(* IEC 61131-3 sources: model-first-plc-agent-ai/results/T3-W-09, 2 files *)

(* ---- a1_code.st ---- *)
FUNCTION_BLOCK TankSequence
VAR_INPUT
    start : BOOL;
    stop : BOOL;
    LSH : BOOL;
    LSHH : BOOL;
    TON_Duration : TIME;
    TOF_Duration : TIME;
END_VAR
VAR_OUTPUT
    fill_valve : BOOL;
    discharge_valve : BOOL;
END_VAR
VAR
    active_state : INT := 0;
    filling_active : BOOL;
    ton_q : BOOL;
    tof_q : BOOL;
    fill_timer : TON;
    pause_timer : TOF;
END_VAR

(* Evaluate both timers every scan using the current filling-step activity. *)
filling_active := (active_state = 1);

fill_timer(IN := filling_active, PT := TON_Duration);
pause_timer(IN := filling_active, PT := TOF_Duration);

ton_q := fill_timer.Q;
tof_q := pause_timer.Q;

(* Evaluate transitions from the current situation only. *)
CASE active_state OF
    0:
        IF start AND NOT stop AND NOT LSH AND NOT LSHH THEN
            active_state := 1;
        END_IF;

    1:
        IF stop OR LSH OR LSHH THEN
            active_state := 0;
        ELSIF ton_q AND NOT stop AND NOT LSH AND NOT LSHH THEN
            active_state := 2;
        END_IF;

    2:
        IF stop OR LSH OR LSHH THEN
            active_state := 0;
        ELSIF NOT tof_q AND NOT stop AND NOT LSH AND NOT LSHH THEN
            active_state := 1;
        END_IF;

ELSE
    active_state := 0;
END_CASE;

(* Continuous actions of the resulting situation. *)
fill_valve := (active_state = 1);
discharge_valve := FALSE;

END_FUNCTION_BLOCK

PROGRAM Main
VAR
    StartCommand AT %IX100.0 : BOOL;
    StopCommand AT %IX100.1 : BOOL;
    LSH AT %IX100.2 : BOOL;
    LSHH AT %IX100.3 : BOOL;
    FillValve AT %QX100.0 : BOOL;
    DischargeValve AT %QX100.1 : BOOL;
END_VAR
VAR
    (* Configurable example presets. *)
    TON_Duration : TIME := T#5s;
    TOF_Duration : TIME := T#5s;
    initialized : BOOL := FALSE;
    start : BOOL := FALSE;
    start_edge : R_TRIG;
    sequence_runtime : TankSequence;
END_VAR

IF NOT initialized THEN
    FillValve := FALSE;
    DischargeValve := FALSE;
    initialized := TRUE;
END_IF;

start_edge(CLK := StartCommand);
start := start_edge.Q;

sequence_runtime(
    start := start,
    stop := StopCommand,
    LSH := LSH,
    LSHH := LSHH,
    TON_Duration := TON_Duration,
    TOF_Duration := TOF_Duration
);

FillValve := sequence_runtime.fill_valve;
DischargeValve := sequence_runtime.discharge_valve;

END_PROGRAM

(* ---- a2_code.st ---- *)
FUNCTION_BLOCK TankFillingControl
VAR_INPUT
    StartCommand : BOOL;
    StopCommand : BOOL;
    LSH : BOOL;
    LSHH : BOOL;
    TON_Duration : TIME;
    TOF_Duration : TIME;
END_VAR
VAR_OUTPUT
    fill_valve : BOOL;
    discharge_valve : BOOL;
END_VAR
VAR
    ActiveState : INT := 0;
    StartEdge : R_TRIG;
    FillingTimer : TON;
    PauseTimer : TOF;
    start : BOOL;
    stop : BOOL;
    ton_q : BOOL;
    tof_q : BOOL;
    FillingActive : BOOL;
END_VAR

StartEdge(CLK := StartCommand);
start := StartEdge.Q;
stop := StopCommand;

FillingActive := (ActiveState = 1);

FillingTimer(
    IN := FillingActive,
    PT := TON_Duration
);

PauseTimer(
    IN := FillingActive,
    PT := TOF_Duration
);

ton_q := FillingTimer.Q;
tof_q := PauseTimer.Q;

IF stop THEN
    ActiveState := 0;
ELSE
    CASE ActiveState OF
        0:
            IF start AND NOT LSH THEN
                ActiveState := 1;
            END_IF;

        1:
            IF LSH THEN
                ActiveState := 0;
            ELSIF ton_q THEN
                ActiveState := 2;
            END_IF;

        2:
            IF LSH THEN
                ActiveState := 0;
            ELSIF NOT tof_q THEN
                ActiveState := 1;
            END_IF;

        ELSE
            ActiveState := 0;
    END_CASE;
END_IF;

fill_valve := (ActiveState = 1) AND NOT stop;
discharge_valve := FALSE;

(* LSHH is an observation input; the specified GRAFCET defines
   no additional transition or interlock for this signal. *)

END_FUNCTION_BLOCK

PROGRAM Main
VAR
    StartCommand AT %IX100.0 : BOOL;
    StopCommand AT %IX100.1 : BOOL;
    LSH AT %IX100.2 : BOOL;
    LSHH AT %IX100.3 : BOOL;
    FillValve AT %QX100.0 : BOOL;
    DischargeValve AT %QX100.1 : BOOL;
END_VAR
VAR
    TankController : TankFillingControl;
    (* Example presets; configure these for the plant. *)
    TON_Duration : TIME := T#5s;
    TOF_Duration : TIME := T#5s;
END_VAR

TankController(
    StartCommand := StartCommand,
    StopCommand := StopCommand,
    LSH := LSH,
    LSHH := LSHH,
    TON_Duration := TON_Duration,
    TOF_Duration := TOF_Duration
);

FillValve := TankController.fill_valve;
DischargeValve := TankController.discharge_valve;

END_PROGRAM
